// TIA Portal project "000000000000-某某-基于顺序控制的交通灯控制系统设计" (V15)

(* hardware
DEVICE "S7-1200 station_1"  S7-1200 Station
   slot 0: "Rack_0"  S7-1200 Rack  Rack  V1.0
   slot 1: "PLC_1"  CPU 1214C DC/DC/Rly  6ES7 214-1HG40-0XB0  V4.2
*)

// ===== PLC "PLC_1"  CPU 1214C DC/DC/Rly =====

VAR_GLOBAL   // PLC tag table "默认变量表"
   "模式选择" AT %I0.0 : Bool;
   "启动按钮" AT %I0.1 : Bool;
   "停止按钮" AT %I0.2 : Bool;
   "东西红灯" AT %Q0.0 : Bool;
   "东西黄灯" AT %Q0.1 : Bool;
   "东西绿灯" AT %Q0.2 : Bool;
   "南北红灯" AT %Q0.3 : Bool;
   "南北黄灯" AT %Q0.4 : Bool;
   "南北绿灯" AT %Q0.5 : Bool;
   "System_Byte" AT %MB10 : Byte;
   "FirstScan" AT %M10.0 : Bool;
   "DiagStatusUpdate" AT %M10.1 : Bool;
   "AlwaysTRUE" AT %M10.2 : Bool;
   "AlwaysFALSE" AT %M10.3 : Bool;
   "Clock_Byte" AT %MB5 : Byte;
   "Clock_10Hz" AT %M5.0 : Bool;
   "Clock_5Hz" AT %M5.1 : Bool;
   "Clock_2.5Hz" AT %M5.2 : Bool;
   "Clock_2Hz" AT %M5.3 : Bool;
   "Clock_1.25Hz" AT %M5.4 : Bool;
   "Clock_1Hz" AT %M5.5 : Bool;
   "Clock_0.625Hz" AT %M5.6 : Bool;
   "Clock_0.5Hz" AT %M5.7 : Bool;
   "M0.0" AT %M0.0 : Bool;
   "M0.1" AT %M0.1 : Bool;
   "M0.2" AT %M0.2 : Bool;
   "M0.3" AT %M0.3 : Bool;
   "M0.4" AT %M0.4 : Bool;
   "M1.1" AT %M1.1 : Bool;
   "M1.2" AT %M1.2 : Bool;
   "M1.3" AT %M1.3 : Bool;
   "M1.4" AT %M1.4 : Bool;
   "M2.0" AT %M2.0 : Bool;
   "M3.0" AT %M3.0 : Bool;
   "Tag_1" AT %MD10 : Time;
   "Tag_2" AT %MD14 : Time;
   "Tag_3" AT %MD18 : Time;
   "Tag_4" AT %MD22 : Time;
   "Tag_5" AT %MD26 : Time;
   "Tag_6" AT %MD30 : Time;
   "Tag_7" AT %MD34 : Time;
   "Tag_8" AT %MD38 : Time;
END_VAR

// folder: System blocks/Program resources

DATA_BLOCK "东西红灯20S"   // DB1
{ S7_Optimized_Access := 'TRUE' }
AUTHOR : Simatic
FAMILY : IEC
NAME : IEC_TMR
VERSION : 1.0
// stored: InstanceOfName IEC_TIMER
"IEC_TIMER"
BEGIN
END_DATA_BLOCK

DATA_BLOCK "东西绿灯15S"   // DB2
{ S7_Optimized_Access := 'TRUE' }
AUTHOR : Simatic
FAMILY : IEC
NAME : IEC_TMR
VERSION : 1.0
// stored: InstanceOfName IEC_TIMER
"IEC_TIMER"
BEGIN
END_DATA_BLOCK

DATA_BLOCK "东西绿灯闪烁3S"   // DB3
{ S7_Optimized_Access := 'TRUE' }
AUTHOR : Simatic
FAMILY : IEC
NAME : IEC_TMR
VERSION : 1.0
// stored: InstanceOfName IEC_TIMER
"IEC_TIMER"
BEGIN
END_DATA_BLOCK

DATA_BLOCK "东西黄灯2S"   // DB4
{ S7_Optimized_Access := 'TRUE' }
AUTHOR : Simatic
FAMILY : IEC
NAME : IEC_TMR
VERSION : 1.0
// stored: InstanceOfName IEC_TIMER
"IEC_TIMER"
BEGIN
END_DATA_BLOCK

DATA_BLOCK "南北绿灯15S"   // DB5
{ S7_Optimized_Access := 'TRUE' }
AUTHOR : Simatic
FAMILY : IEC
NAME : IEC_TMR
VERSION : 1.0
// stored: InstanceOfName IEC_TIMER
"IEC_TIMER"
BEGIN
END_DATA_BLOCK

DATA_BLOCK "南北绿灯闪烁3S"   // DB6
{ S7_Optimized_Access := 'TRUE' }
AUTHOR : Simatic
FAMILY : IEC
NAME : IEC_TMR
VERSION : 1.0
// stored: InstanceOfName IEC_TIMER
"IEC_TIMER"
BEGIN
END_DATA_BLOCK

DATA_BLOCK "南北黄灯闪烁2S"   // DB7
{ S7_Optimized_Access := 'TRUE' }
AUTHOR : Simatic
FAMILY : IEC
NAME : IEC_TMR
VERSION : 1.0
// stored: InstanceOfName IEC_TIMER
"IEC_TIMER"
BEGIN
END_DATA_BLOCK

DATA_BLOCK "南北红灯20S"   // DB8
{ S7_Optimized_Access := 'TRUE' }
AUTHOR : Simatic
FAMILY : IEC
NAME : IEC_TMR
VERSION : 1.0
// stored: InstanceOfName IEC_TIMER
"IEC_TIMER"
BEGIN
END_DATA_BLOCK

// folder: (top level)

ORGANIZATION_BLOCK "Main"   // OB1, LAD, ProgramCycle
TITLE = "Main Program Sweep (Cycle)"
{ S7_Optimized_Access := 'TRUE' }
VERSION : 0.1
   VAR_INPUT
      Initial_Call : Bool;   // Initial call of this OB
      Remanence : Bool;   // =True, if remanent data are available
   END_VAR
   VAR_TEMP   // added for the SCL form of the ladder/FBD networks
      _w1 : Bool;
      _w2 : Bool;
      _w3 : Bool;
      _w4 : Bool;
      _w5 : Bool;
   END_VAR
BEGIN

REGION Network 1: 开始
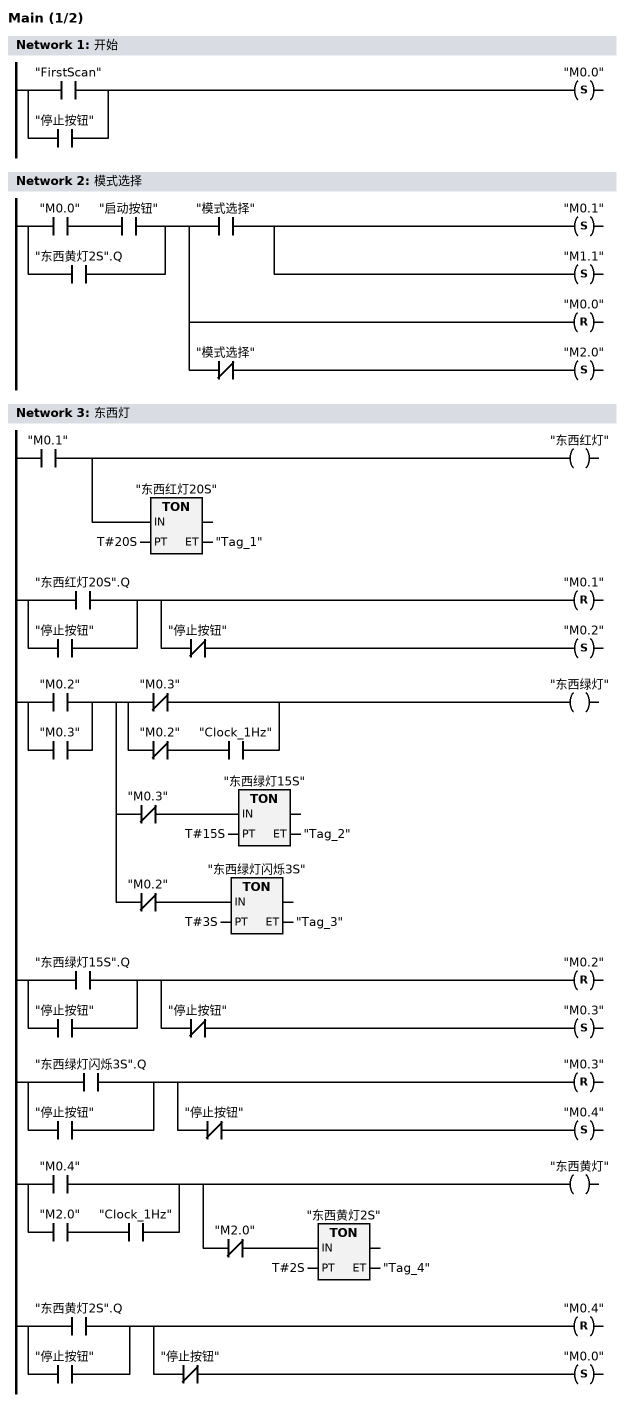
   RUNG wire#powerrail
      Contact( "FirstScan" )
      wire#w1
      S_Coil( "M0.0" )
   END_RUNG
   RUNG wire#powerrail
      Contact( "停止按钮" )
   END_RUNG wire#w1
   // the same network as SCL:
   IF "FirstScan" OR "停止按钮" THEN "M0.0" := TRUE; END_IF;
END_REGION

REGION Network 2: 模式选择
   RUNG wire#powerrail
      Contact( "M0.0" )
      Contact( "启动按钮" )
      wire#w1
      Contact( "模式选择" )
      wire#w2
      S_Coil( "M0.1" )
   END_RUNG
   RUNG wire#powerrail
      Contact( "东西黄灯2S".Q )
   END_RUNG wire#w1
   RUNG wire#w2
      S_Coil( "M1.1" )
   END_RUNG
   RUNG wire#w1
      R_Coil( "M0.0" )
   END_RUNG
   RUNG wire#w1
      I_Contact( "模式选择" )
      S_Coil( "M2.0" )
   END_RUNG
   // the same network as SCL:
   #_w1 := ("M0.0" AND "启动按钮") OR "东西黄灯2S".Q;
   IF #_w1 AND "模式选择" THEN
       "M0.1" := TRUE;
       "M1.1" := TRUE;
   END_IF;
   IF #_w1 THEN "M0.0" := FALSE; END_IF;
   IF #_w1 AND NOT "模式选择" THEN "M2.0" := TRUE; END_IF;
END_REGION

REGION Network 3: 东西灯
   "东西红灯" := "M0.1";
   "东西红灯20S".TON(IN := "M0.1", PT := T#20S, ET => "Tag_1");
   #_w1 := "东西红灯20S".Q OR "停止按钮";
   IF #_w1 THEN "M0.1" := FALSE; END_IF;
   IF #_w1 AND NOT "停止按钮" THEN "M0.2" := TRUE; END_IF;
   #_w2 := "M0.2" OR "M0.3";
   "东西绿灯" := #_w2 AND (NOT "M0.3" OR (NOT "M0.2" AND "Clock_1Hz"));
   "东西绿灯15S".TON(IN := #_w2 AND NOT "M0.3", PT := T#15S, ET => "Tag_2");
   "东西绿灯闪烁3S".TON(IN := #_w2 AND NOT "M0.2", PT := T#3S, ET => "Tag_3");
   #_w3 := "东西绿灯15S".Q OR "停止按钮";
   IF #_w3 THEN "M0.2" := FALSE; END_IF;
   IF #_w3 AND NOT "停止按钮" THEN "M0.3" := TRUE; END_IF;
   #_w4 := "东西绿灯闪烁3S".Q OR "停止按钮";
   IF #_w4 THEN "M0.3" := FALSE; END_IF;
   IF #_w4 AND NOT "停止按钮" THEN "M0.4" := TRUE; END_IF;
   "东西黄灯" := "M0.4" OR ("M2.0" AND "Clock_1Hz");
   "东西黄灯2S".TON(IN := "东西黄灯" AND NOT "M2.0", PT := T#2S, ET => "Tag_4");
   #_w5 := "东西黄灯2S".Q OR "停止按钮";
   IF #_w5 THEN "M0.4" := FALSE; END_IF;
   IF #_w5 AND NOT "停止按钮" THEN "M0.0" := TRUE; END_IF;
END_REGION

REGION Network 4: 南北灯
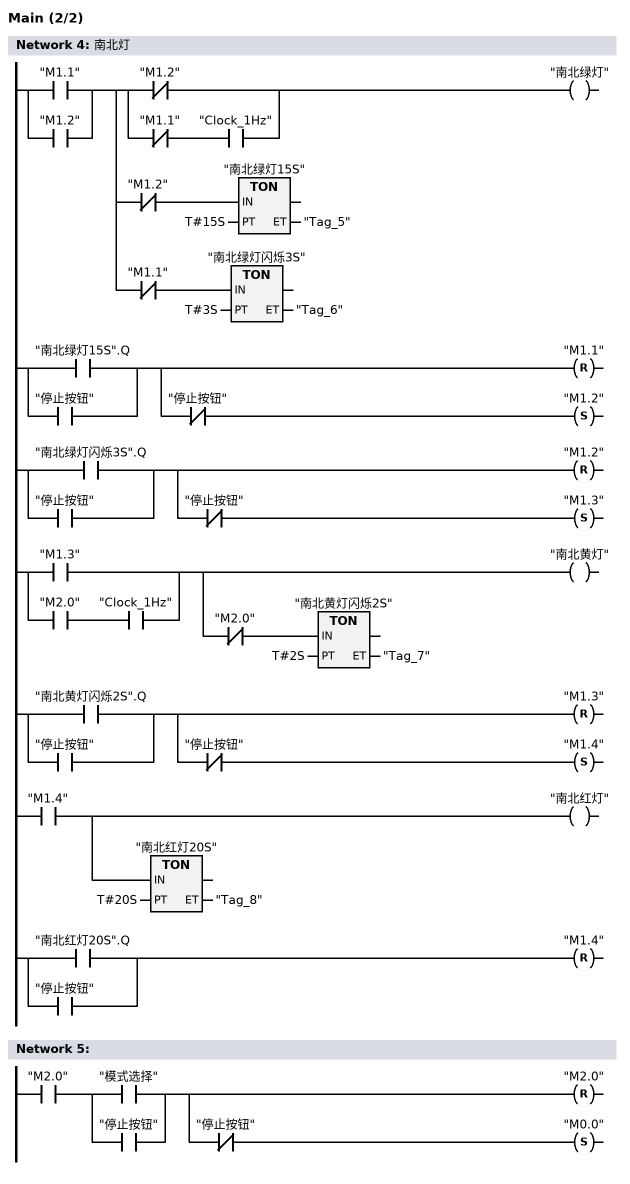
   #_w1 := "M1.1" OR "M1.2";
   "南北绿灯" := #_w1 AND (NOT "M1.2" OR (NOT "M1.1" AND "Clock_1Hz"));
   "南北绿灯15S".TON(IN := #_w1 AND NOT "M1.2", PT := T#15S, ET => "Tag_5");
   "南北绿灯闪烁3S".TON(IN := #_w1 AND NOT "M1.1", PT := T#3S, ET => "Tag_6");
   #_w2 := "南北绿灯15S".Q OR "停止按钮";
   IF #_w2 THEN "M1.1" := FALSE; END_IF;
   IF #_w2 AND NOT "停止按钮" THEN "M1.2" := TRUE; END_IF;
   #_w3 := "南北绿灯闪烁3S".Q OR "停止按钮";
   IF #_w3 THEN "M1.2" := FALSE; END_IF;
   IF #_w3 AND NOT "停止按钮" THEN "M1.3" := TRUE; END_IF;
   "南北黄灯" := "M1.3" OR ("M2.0" AND "Clock_1Hz");
   "南北黄灯闪烁2S".TON(IN := "南北黄灯" AND NOT "M2.0", PT := T#2S, ET => "Tag_7");
   #_w4 := "南北黄灯闪烁2S".Q OR "停止按钮";
   IF #_w4 THEN "M1.3" := FALSE; END_IF;
   IF #_w4 AND NOT "停止按钮" THEN "M1.4" := TRUE; END_IF;
   "南北红灯" := "M1.4";
   "南北红灯20S".TON(IN := "M1.4", PT := T#20S, ET => "Tag_8");
   IF "南北红灯20S".Q OR "停止按钮" THEN "M1.4" := FALSE; END_IF;
END_REGION

REGION Network 5
   RUNG wire#powerrail
      Contact( "M2.0" )
      wire#w1
      Contact( "模式选择" )
      wire#w2
      R_Coil( "M2.0" )
   END_RUNG
   RUNG wire#w1
      Contact( "停止按钮" )
   END_RUNG wire#w2
   RUNG wire#w2
      I_Contact( "停止按钮" )
      S_Coil( "M0.0" )
   END_RUNG
   // the same network as SCL:
   #_w1 := "M2.0" AND ("模式选择" OR "停止按钮");
   IF #_w1 THEN "M2.0" := FALSE; END_IF;
   IF #_w1 AND NOT "停止按钮" THEN "M0.0" := TRUE; END_IF;
END_REGION
END_ORGANIZATION_BLOCK